Fanuc KAREL source: KC00056.KL

PROGRAM KC00056
%NOLOCKGROUP
%ENVIRONMENT DEBUG
VAR
  I: INTEGER
  J: INTEGER
  K: INTEGER
  R: REAL
  B: BOOLEAN
  S: STRING[80]
  T: STRING[80]
  P: PATH
  Q: PATH
  AI: ARRAY[8] OF INTEGER
  AB: ARRAY[244] OF BYTE
BEGIN
  SET_DEBUG(B)
END KC00056
